FUNCTION F_ModDW : DWORD
(*
Modulo function for double word numbers (dividend mod divisor).

Constructor: 		Patryk Panylo
Company:		E. Riexinger GmbH
Date:			20.01.2014
Version:			1.00

Date:			Revision:		Who:				Comment
dd.mm.yyyy		x.xx			Initials			comment

*)
VAR_INPUT
	dwDividend						:DWORD;
	dwDivisor						:DWORD;
END_VAR
VAR
END_VAR


F_MODDW := dwDivisor;

IF dwDivisor <> 0 
THEN
	F_MODDW := dwDividend MOD dwDivisor;
END_IF;

END_FUNCTION

(* stored: Version 1.1.0.1, ProductVersion 3.1.4024.15
   POU F_ModDW: Id {13cd23a6-ba05-46db-baff-b193e3e1e2e5}, SpecialFunc None *)
